Fanuc KAREL source: kb00039.KL

-- PROVISIONAL review KL for V770-1; original PC SHA256 d54cb02556c7282684fb767eb52990cfd3cd15231634288164a57cb32a161f39
-- Incomplete behavior may be omitted. Consult companion uncertainty JSON. Do not deploy.
PROGRAM KB00039
%NOLOCKGROUP
BEGIN
  -- UNRESOLVED_PC offsets 5-14; opcodes 3F,75
  -- UNRESOLVED_PC offsets 19-26; opcodes 9D,23
  -- UNRESOLVED_PC offsets 31-55; opcodes 27,22,2A,22,22,31
  -- UNRESOLVED_PC offsets 60-64; opcodes 7F
END KB00039
